(*
SPDX-License-Identifier: MIT
License: https://opensource.org/license/mit
*)

(*!
<summary>Owns a timer-delay test as a static group.</summary>
<description>
Owns persistent child storage and fixed parent associations. Use in one task without reentry.
Children is borrowed and must not be modified by application code. Constructor callbacks are not used.
</description>
*)

{attribute 'no_assign'}
{attribute 'no_explicit_call' := 'do not call this function block directly'}
FUNCTION_BLOCK TimingTestGroup EXTENDS TOF_Testing.TestGroup<1>
VAR_STAT
	//! <summary>Class name shared by all instances of this function block.</summary>
	{attribute 'hide'}
	_ClassName : STRING := __POUNAME();
END_VAR
VAR
	_Timer : TimerDelayTest(name := "Timer delay", parent := THIS^);

	_Children : ARRAY [0.._ChildCount - 1] OF TOF_Testing.ITestElement :=
	[
		_Timer
	];
END_VAR

//! <summary>Borrows the fixed array of this concrete group; do not modify it.</summary>
{attribute 'monitoring' := 'call'}
PROPERTY Children : REFERENCE TO ARRAY [0.._ChildCount - 1] OF TOF_Testing.ITestElement
GET
Children REF= _Children;
END_GET
END_PROPERTY

//! <summary>Borrows the concrete class name for the lifetime of this instance; callers must not modify it.</summary>
{attribute 'monitoring' := 'call'}
PROPERTY ClassName : REFERENCE TO STRING
GET
ClassName REF= _ClassName;
END_GET
END_PROPERTY

//! <summary>Borrows the compiler-initialized namespace; callers must not modify the returned reference.</summary>
{attribute 'monitoring' := 'call'}
PROPERTY NamespaceName : REFERENCE TO STRING
GET
NamespaceName REF= CurrentNamespace.Name;
END_GET
END_PROPERTY

//! <summary>Reports the complete concrete instance size, excluding separately allocated storage.</summary>
{attribute 'monitoring' := 'call'}
PROPERTY SelfSize : ULINT
GET
SelfSize := XSIZEOF(THIS^);
END_GET
END_PROPERTY

END_FUNCTION_BLOCK

(* stored: Version 1.1.0.1
   POU TimingTestGroup: Id {34539cb8-6b6e-4ea1-b7e6-d4e6b19474ee}, SpecialFunc None
   Property Children: Id {c8b52158-bb93-4786-9d76-fa1c263f917e}
   Get Get: Id {08e1ae17-0f95-48b2-baac-a2797cb32562}
   Property ClassName: Id {55b5ff7b-61ba-4422-b80d-e77b9f6b1006}
   Get Get: Id {b9f63e33-f26e-47ff-bad3-67e2df9eff89}
   Property NamespaceName: Id {62dd84d1-718e-4ecf-96b6-47c0041b7513}
   Get Get: Id {bc3ba1a4-ed59-417a-90b4-00654202621c}
   Property SelfSize: Id {18b4faf7-49f5-4a54-97ef-cad8c0a1272a}
   Get Get: Id {71891571-1736-4071-816b-df3f352603ca} *)
